FUNCTION_BLOCK SKILL_FailMerge (* Joins two failure events (with their error codes) into one, because a data input can only be wired once. Technical: Merges two failure events with their error codes into one *)
  (* Standard: 61499-2 *)
  (* Version 0.1, 2026-09-28, Project contributors, AAU Smart Production Lab *)
  PACKAGE modlib;
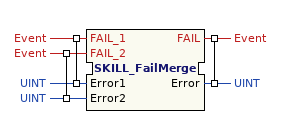
  EVENT_INPUT
    FAIL_1 WITH Error1; (* A step failed (Error1) *)
    FAIL_2 WITH Error2; (* A step failed (Error2) *)
  END_EVENT
  EVENT_OUTPUT
    FAIL WITH Error; (* One of them failed (Error) *)
  END_EVENT
  VAR_INPUT
    Error1 : UINT; (* Error code of the first *)
    Error2 : UINT; (* Error code of the second *)
  END_VAR
  VAR_OUTPUT
    Error : UINT; (* Error code of the one that failed *)
  END_VAR
  EC_STATES
    FAIL_1 : FAIL_1 -> FAIL;
    FAIL_2 : FAIL_2 -> FAIL;
  END_STATES
  ALGORITHM FAIL_1 IN ST:
Error := Error1;
  END_ALGORITHM
  ALGORITHM FAIL_2 IN ST:
Error := Error2;
  END_ALGORITHM
END_FUNCTION_BLOCK
